FUNCTION_BLOCK BATCH_FILLING (* Migrated from IEC 61131-3 ST *)
  (* Standard: 61499-2 *)
  (* Version 1.0, 2026-11-06, st2fb *)
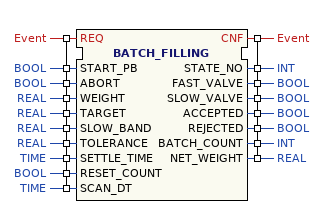
  EVENT_INPUT
    REQ WITH START_PB, ABORT, WEIGHT, TARGET, SLOW_BAND, TOLERANCE, SETTLE_TIME, RESET_COUNT, SCAN_DT;
  END_EVENT
  EVENT_OUTPUT
    CNF WITH STATE_NO, FAST_VALVE, SLOW_VALVE, ACCEPTED, REJECTED, BATCH_COUNT, NET_WEIGHT;
  END_EVENT
  VAR_INPUT
    START_PB : BOOL;
    ABORT : BOOL;
    WEIGHT : REAL;
    TARGET : REAL;
    SLOW_BAND : REAL;
    TOLERANCE : REAL;
    SETTLE_TIME : TIME;
    RESET_COUNT : BOOL;
    SCAN_DT : TIME;
  END_VAR
  VAR_OUTPUT
    STATE_NO : INT;
    FAST_VALVE : BOOL;
    SLOW_VALVE : BOOL;
    ACCEPTED : BOOL;
    REJECTED : BOOL;
    BATCH_COUNT : INT;
    NET_WEIGHT : REAL;
  END_VAR
  VAR
    TARE : REAL;
    COUNT_PULSE : BOOL;
    ST2FB_NOW : TIME := T#0s;
    START_EDGE_CLK : BOOL;
    START_EDGE_Q : BOOL;
    START_EDGE_M : BOOL;
    SETTLE_TIMER_IN : BOOL;
    SETTLE_TIMER_PT : TIME;
    SETTLE_TIMER_Q : BOOL;
    SETTLE_TIMER_ET : TIME;
    SETTLE_TIMER_STATE : INT;
    SETTLE_TIMER_PREV_IN : BOOL;
    SETTLE_TIMER_START_TIME : TIME;
    COUNTER_CU : BOOL;
    COUNTER_R : BOOL;
    COUNTER_PV : INT;
    COUNTER_Q : BOOL;
    COUNTER_CV : INT;
    COUNTER_CU_T_Q : BOOL;
    COUNTER_CU_T_M : BOOL;
  END_VAR
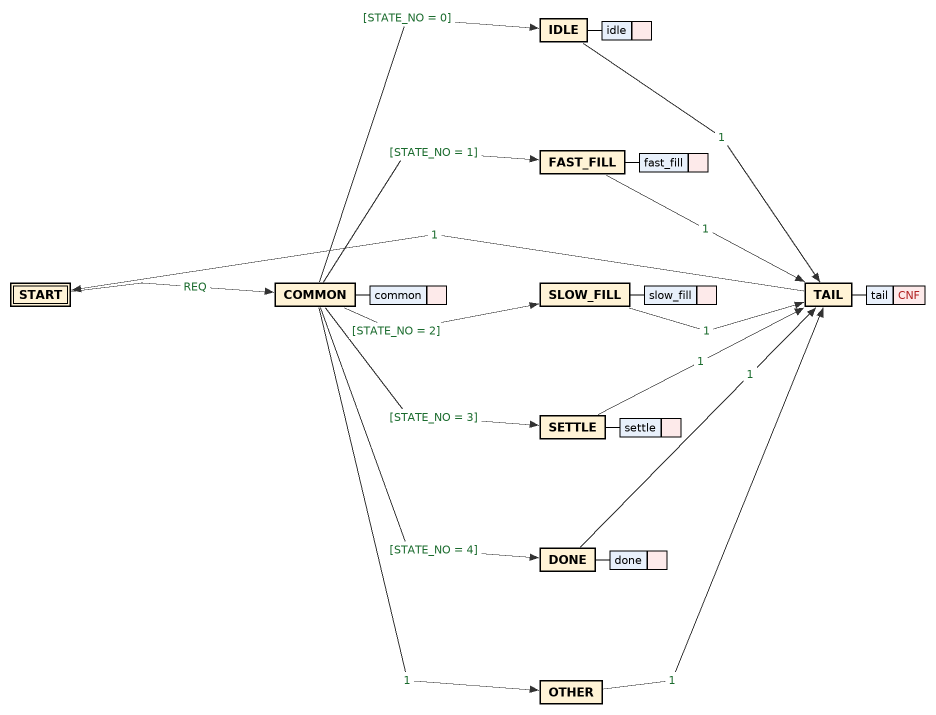
  EC_STATES
    START;
    COMMON : common;
    IDLE : idle;
    FAST_FILL : fast_fill;
    SLOW_FILL : slow_fill;
    SETTLE : settle;
    DONE : done;
    OTHER;
    TAIL : tail -> CNF;
  END_STATES
  EC_TRANSITIONS
    START TO COMMON := REQ;
    COMMON TO IDLE := [STATE_NO = 0];
    COMMON TO FAST_FILL := [STATE_NO = 1];
    COMMON TO SLOW_FILL := [STATE_NO = 2];
    COMMON TO SETTLE := [STATE_NO = 3];
    COMMON TO DONE := [STATE_NO = 4];
    COMMON TO OTHER := 1;
    IDLE TO TAIL := 1;
    FAST_FILL TO TAIL := 1;
    SLOW_FILL TO TAIL := 1;
    SETTLE TO TAIL := 1;
    DONE TO TAIL := 1;
    OTHER TO TAIL := 1;
    TAIL TO START := 1;
  END_TRANSITIONS
  ALGORITHM common IN ST:
ST2FB_NOW := ST2FB_NOW + SCAN_DT;
START_EDGE_CLK := START_PB;
START_EDGE_Q := START_EDGE_CLK AND NOT START_EDGE_M;
START_EDGE_M := START_EDGE_CLK;
NET_WEIGHT := WEIGHT - TARE;
FAST_VALVE := FALSE;
SLOW_VALVE := FALSE;
COUNT_PULSE := FALSE;
IF ABORT THEN
  STATE_NO := 0;
  ACCEPTED := FALSE;
  REJECTED := FALSE;
END_IF;
  END_ALGORITHM
  ALGORITHM idle IN ST:
IF START_EDGE_Q AND NOT ABORT THEN
  TARE := WEIGHT;
  NET_WEIGHT := 0.0;
  ACCEPTED := FALSE;
  REJECTED := FALSE;
  STATE_NO := 1;
END_IF;
  END_ALGORITHM
  ALGORITHM fast_fill IN ST:
FAST_VALVE := TRUE;
SLOW_VALVE := TRUE;
IF NET_WEIGHT >= TARGET - SLOW_BAND THEN
  STATE_NO := 2;
END_IF;
  END_ALGORITHM
  ALGORITHM slow_fill IN ST:
SLOW_VALVE := TRUE;
IF NET_WEIGHT >= TARGET THEN
  STATE_NO := 3;
END_IF;
  END_ALGORITHM
  ALGORITHM settle IN ST:
IF SETTLE_TIMER_Q THEN
  IF (NET_WEIGHT >= TARGET - TOLERANCE) AND (NET_WEIGHT <= TARGET + TOLERANCE) THEN
    ACCEPTED := TRUE;
    COUNT_PULSE := TRUE;
  ELSE
    REJECTED := TRUE;
  END_IF;
  STATE_NO := 4;
END_IF;
  END_ALGORITHM
  ALGORITHM done IN ST:
IF START_EDGE_Q THEN
  TARE := WEIGHT;
  NET_WEIGHT := 0.0;
  ACCEPTED := FALSE;
  REJECTED := FALSE;
  STATE_NO := 1;
END_IF;
  END_ALGORITHM
  ALGORITHM tail IN ST:
SETTLE_TIMER_IN := STATE_NO = 3;
SETTLE_TIMER_PT := SETTLE_TIME;
IF (SETTLE_TIMER_STATE = 0) AND NOT SETTLE_TIMER_PREV_IN AND SETTLE_TIMER_IN THEN
  SETTLE_TIMER_STATE := 1;
  SETTLE_TIMER_Q := FALSE;
  SETTLE_TIMER_START_TIME := ST2FB_NOW;
ELSE
  IF NOT SETTLE_TIMER_IN THEN
    SETTLE_TIMER_ET := T#0s;
    SETTLE_TIMER_Q := FALSE;
    SETTLE_TIMER_STATE := 0;
  ELSIF SETTLE_TIMER_STATE = 1 THEN
    IF SETTLE_TIMER_START_TIME + SETTLE_TIMER_PT <= ST2FB_NOW THEN
      SETTLE_TIMER_STATE := 2;
      SETTLE_TIMER_Q := TRUE;
      SETTLE_TIMER_ET := SETTLE_TIMER_PT;
    ELSE
      SETTLE_TIMER_ET := ST2FB_NOW - SETTLE_TIMER_START_TIME;
    END_IF;
  END_IF;
END_IF;
SETTLE_TIMER_PREV_IN := SETTLE_TIMER_IN;
COUNTER_CU := COUNT_PULSE;
COUNTER_R := RESET_COUNT;
COUNTER_PV := 1000;
COUNTER_CU_T_Q := COUNTER_CU AND NOT COUNTER_CU_T_M;
COUNTER_CU_T_M := COUNTER_CU;
IF COUNTER_R THEN
  COUNTER_CV := 0;
ELSIF COUNTER_CU_T_Q AND (COUNTER_CV < COUNTER_PV) THEN
  COUNTER_CV := COUNTER_CV + 1;
END_IF;
COUNTER_Q := COUNTER_CV >= COUNTER_PV;
BATCH_COUNT := COUNTER_CV;
  END_ALGORITHM
END_FUNCTION_BLOCK
